(* IEC 61131-3 sources: STAR-PLC-Agent/results/raw/codex_matrix_resume_20261114/codex_deepseek/PUB002/functional/attempt_0001, 1 file *)

(* ---- test_program.st ---- *)
PROGRAM PLC_PRG
VAR
 BenchStep : UDINT := 0;
 BenchCalls : UDINT := 0;
 BenchDone : BOOL := FALSE;
 BenchUut0 : FB_Task;
 BenchUut1 : FB_Task;
 BenchUut2 : FB_Task;
 BenchUut3 : FB_Task;
 BenchUut4 : FB_Task;
 BenchUut5 : FB_Task;
 BenchUut6 : FB_Task;
 TraceIn_value : ARRAY[0..38] OF DWORD;
 TraceOut_hasChanged : ARRAY[0..38] OF BOOL;
 TraceOut_hasRisingEdges : ARRAY[0..38] OF BOOL;
 TraceOut_risingBits : ARRAY[0..38] OF DWORD;
 TraceOut_noOfRisingBits : ARRAY[0..38] OF USINT;
 TraceOut_hasFallingEdges : ARRAY[0..38] OF BOOL;
 TraceOut_fallingBits : ARRAY[0..38] OF DWORD;
 TraceOut_noOfFallingBits : ARRAY[0..38] OF USINT;
END_VAR

IF NOT BenchDone THEN
 CASE BenchStep OF
 0:
   BenchUut0.value := DWORD#0;
   TraceIn_value[0] := BenchUut0.value;
   BenchUut0();
   TraceOut_hasChanged[0] := BenchUut0.hasChanged;
   TraceOut_hasRisingEdges[0] := BenchUut0.hasRisingEdges;
   TraceOut_risingBits[0] := BenchUut0.risingBits;
   TraceOut_noOfRisingBits[0] := BenchUut0.noOfRisingBits;
   TraceOut_hasFallingEdges[0] := BenchUut0.hasFallingEdges;
   TraceOut_fallingBits[0] := BenchUut0.fallingBits;
   TraceOut_noOfFallingBits[0] := BenchUut0.noOfFallingBits;
   BenchCalls := BenchCalls + 1;
 1:
   BenchUut0.value := DWORD#1;
   TraceIn_value[1] := BenchUut0.value;
   BenchUut0();
   TraceOut_hasChanged[1] := BenchUut0.hasChanged;
   TraceOut_hasRisingEdges[1] := BenchUut0.hasRisingEdges;
   TraceOut_risingBits[1] := BenchUut0.risingBits;
   TraceOut_noOfRisingBits[1] := BenchUut0.noOfRisingBits;
   TraceOut_hasFallingEdges[1] := BenchUut0.hasFallingEdges;
   TraceOut_fallingBits[1] := BenchUut0.fallingBits;
   TraceOut_noOfFallingBits[1] := BenchUut0.noOfFallingBits;
   BenchCalls := BenchCalls + 1;
 2:
   BenchUut0.value := DWORD#1;
   TraceIn_value[2] := BenchUut0.value;
   BenchUut0();
   TraceOut_hasChanged[2] := BenchUut0.hasChanged;
   TraceOut_hasRisingEdges[2] := BenchUut0.hasRisingEdges;
   TraceOut_risingBits[2] := BenchUut0.risingBits;
   TraceOut_noOfRisingBits[2] := BenchUut0.noOfRisingBits;
   TraceOut_hasFallingEdges[2] := BenchUut0.hasFallingEdges;
   TraceOut_fallingBits[2] := BenchUut0.fallingBits;
   TraceOut_noOfFallingBits[2] := BenchUut0.noOfFallingBits;
   BenchCalls := BenchCalls + 1;
 3:
   BenchUut0.value := DWORD#3;
   TraceIn_value[3] := BenchUut0.value;
   BenchUut0();
   TraceOut_hasChanged[3] := BenchUut0.hasChanged;
   TraceOut_hasRisingEdges[3] := BenchUut0.hasRisingEdges;
   TraceOut_risingBits[3] := BenchUut0.risingBits;
   TraceOut_noOfRisingBits[3] := BenchUut0.noOfRisingBits;
   TraceOut_hasFallingEdges[3] := BenchUut0.hasFallingEdges;
   TraceOut_fallingBits[3] := BenchUut0.fallingBits;
   TraceOut_noOfFallingBits[3] := BenchUut0.noOfFallingBits;
   BenchCalls := BenchCalls + 1;
 4:
   BenchUut0.value := DWORD#2;
   TraceIn_value[4] := BenchUut0.value;
   BenchUut0();
   TraceOut_hasChanged[4] := BenchUut0.hasChanged;
   TraceOut_hasRisingEdges[4] := BenchUut0.hasRisingEdges;
   TraceOut_risingBits[4] := BenchUut0.risingBits;
   TraceOut_noOfRisingBits[4] := BenchUut0.noOfRisingBits;
   TraceOut_hasFallingEdges[4] := BenchUut0.hasFallingEdges;
   TraceOut_fallingBits[4] := BenchUut0.fallingBits;
   TraceOut_noOfFallingBits[4] := BenchUut0.noOfFallingBits;
   BenchCalls := BenchCalls + 1;
 5:
   BenchUut0.value := DWORD#0;
   TraceIn_value[5] := BenchUut0.value;
   BenchUut0();
   TraceOut_hasChanged[5] := BenchUut0.hasChanged;
   TraceOut_hasRisingEdges[5] := BenchUut0.hasRisingEdges;
   TraceOut_risingBits[5] := BenchUut0.risingBits;
   TraceOut_noOfRisingBits[5] := BenchUut0.noOfRisingBits;
   TraceOut_hasFallingEdges[5] := BenchUut0.hasFallingEdges;
   TraceOut_fallingBits[5] := BenchUut0.fallingBits;
   TraceOut_noOfFallingBits[5] := BenchUut0.noOfFallingBits;
   BenchCalls := BenchCalls + 1;
 6:
   BenchUut0.value := DWORD#4294967295;
   TraceIn_value[6] := BenchUut0.value;
   BenchUut0();
   TraceOut_hasChanged[6] := BenchUut0.hasChanged;
   TraceOut_hasRisingEdges[6] := BenchUut0.hasRisingEdges;
   TraceOut_risingBits[6] := BenchUut0.risingBits;
   TraceOut_noOfRisingBits[6] := BenchUut0.noOfRisingBits;
   TraceOut_hasFallingEdges[6] := BenchUut0.hasFallingEdges;
   TraceOut_fallingBits[6] := BenchUut0.fallingBits;
   TraceOut_noOfFallingBits[6] := BenchUut0.noOfFallingBits;
   BenchCalls := BenchCalls + 1;
 7:
   BenchUut0.value := DWORD#0;
   TraceIn_value[7] := BenchUut0.value;
   BenchUut0();
   TraceOut_hasChanged[7] := BenchUut0.hasChanged;
   TraceOut_hasRisingEdges[7] := BenchUut0.hasRisingEdges;
   TraceOut_risingBits[7] := BenchUut0.risingBits;
   TraceOut_noOfRisingBits[7] := BenchUut0.noOfRisingBits;
   TraceOut_hasFallingEdges[7] := BenchUut0.hasFallingEdges;
   TraceOut_fallingBits[7] := BenchUut0.fallingBits;
   TraceOut_noOfFallingBits[7] := BenchUut0.noOfFallingBits;
   BenchCalls := BenchCalls + 1;
 8:
   BenchUut0.value := DWORD#2147483648;
   TraceIn_value[8] := BenchUut0.value;
   BenchUut0();
   TraceOut_hasChanged[8] := BenchUut0.hasChanged;
   TraceOut_hasRisingEdges[8] := BenchUut0.hasRisingEdges;
   TraceOut_risingBits[8] := BenchUut0.risingBits;
   TraceOut_noOfRisingBits[8] := BenchUut0.noOfRisingBits;
   TraceOut_hasFallingEdges[8] := BenchUut0.hasFallingEdges;
   TraceOut_fallingBits[8] := BenchUut0.fallingBits;
   TraceOut_noOfFallingBits[8] := BenchUut0.noOfFallingBits;
   BenchCalls := BenchCalls + 1;
 9:
   BenchUut0.value := DWORD#2147483647;
   TraceIn_value[9] := BenchUut0.value;
   BenchUut0();
   TraceOut_hasChanged[9] := BenchUut0.hasChanged;
   TraceOut_hasRisingEdges[9] := BenchUut0.hasRisingEdges;
   TraceOut_risingBits[9] := BenchUut0.risingBits;
   TraceOut_noOfRisingBits[9] := BenchUut0.noOfRisingBits;
   TraceOut_hasFallingEdges[9] := BenchUut0.hasFallingEdges;
   TraceOut_fallingBits[9] := BenchUut0.fallingBits;
   TraceOut_noOfFallingBits[9] := BenchUut0.noOfFallingBits;
   BenchCalls := BenchCalls + 1;
 10:
   BenchUut1.value := DWORD#4294967295;
   TraceIn_value[10] := BenchUut1.value;
   BenchUut1();
   TraceOut_hasChanged[10] := BenchUut1.hasChanged;
   TraceOut_hasRisingEdges[10] := BenchUut1.hasRisingEdges;
   TraceOut_risingBits[10] := BenchUut1.risingBits;
   TraceOut_noOfRisingBits[10] := BenchUut1.noOfRisingBits;
   TraceOut_hasFallingEdges[10] := BenchUut1.hasFallingEdges;
   TraceOut_fallingBits[10] := BenchUut1.fallingBits;
   TraceOut_noOfFallingBits[10] := BenchUut1.noOfFallingBits;
   BenchCalls := BenchCalls + 1;
 11:
   BenchUut1.value := DWORD#4294967295;
   TraceIn_value[11] := BenchUut1.value;
   BenchUut1();
   TraceOut_hasChanged[11] := BenchUut1.hasChanged;
   TraceOut_hasRisingEdges[11] := BenchUut1.hasRisingEdges;
   TraceOut_risingBits[11] := BenchUut1.risingBits;
   TraceOut_noOfRisingBits[11] := BenchUut1.noOfRisingBits;
   TraceOut_hasFallingEdges[11] := BenchUut1.hasFallingEdges;
   TraceOut_fallingBits[11] := BenchUut1.fallingBits;
   TraceOut_noOfFallingBits[11] := BenchUut1.noOfFallingBits;
   BenchCalls := BenchCalls + 1;
 12:
   BenchUut2.value := DWORD#2863311530;
   TraceIn_value[12] := BenchUut2.value;
   BenchUut2();
   TraceOut_hasChanged[12] := BenchUut2.hasChanged;
   TraceOut_hasRisingEdges[12] := BenchUut2.hasRisingEdges;
   TraceOut_risingBits[12] := BenchUut2.risingBits;
   TraceOut_noOfRisingBits[12] := BenchUut2.noOfRisingBits;
   TraceOut_hasFallingEdges[12] := BenchUut2.hasFallingEdges;
   TraceOut_fallingBits[12] := BenchUut2.fallingBits;
   TraceOut_noOfFallingBits[12] := BenchUut2.noOfFallingBits;
   BenchCalls := BenchCalls + 1;
 13:
   BenchUut2.value := DWORD#1431655765;
   TraceIn_value[13] := BenchUut2.value;
   BenchUut2();
   TraceOut_hasChanged[13] := BenchUut2.hasChanged;
   TraceOut_hasRisingEdges[13] := BenchUut2.hasRisingEdges;
   TraceOut_risingBits[13] := BenchUut2.risingBits;
   TraceOut_noOfRisingBits[13] := BenchUut2.noOfRisingBits;
   TraceOut_hasFallingEdges[13] := BenchUut2.hasFallingEdges;
   TraceOut_fallingBits[13] := BenchUut2.fallingBits;
   TraceOut_noOfFallingBits[13] := BenchUut2.noOfFallingBits;
   BenchCalls := BenchCalls + 1;
 14:
   BenchUut3.value := DWORD#983295;
   TraceIn_value[14] := BenchUut3.value;
   BenchUut3();
   TraceOut_hasChanged[14] := BenchUut3.hasChanged;
   TraceOut_hasRisingEdges[14] := BenchUut3.hasRisingEdges;
   TraceOut_risingBits[14] := BenchUut3.risingBits;
   TraceOut_noOfRisingBits[14] := BenchUut3.noOfRisingBits;
   TraceOut_hasFallingEdges[14] := BenchUut3.hasFallingEdges;
   TraceOut_fallingBits[14] := BenchUut3.fallingBits;
   TraceOut_noOfFallingBits[14] := BenchUut3.noOfFallingBits;
   BenchCalls := BenchCalls + 1;
 15:
   BenchUut3.value := DWORD#16715520;
   TraceIn_value[15] := BenchUut3.value;
   BenchUut3();
   TraceOut_hasChanged[15] := BenchUut3.hasChanged;
   TraceOut_hasRisingEdges[15] := BenchUut3.hasRisingEdges;
   TraceOut_risingBits[15] := BenchUut3.risingBits;
   TraceOut_noOfRisingBits[15] := BenchUut3.noOfRisingBits;
   TraceOut_hasFallingEdges[15] := BenchUut3.hasFallingEdges;
   TraceOut_fallingBits[15] := BenchUut3.fallingBits;
   TraceOut_noOfFallingBits[15] := BenchUut3.noOfFallingBits;
   BenchCalls := BenchCalls + 1;
 16:
   BenchUut3.value := DWORD#16715520;
   TraceIn_value[16] := BenchUut3.value;
   BenchUut3();
   TraceOut_hasChanged[16] := BenchUut3.hasChanged;
   TraceOut_hasRisingEdges[16] := BenchUut3.hasRisingEdges;
   TraceOut_risingBits[16] := BenchUut3.risingBits;
   TraceOut_noOfRisingBits[16] := BenchUut3.noOfRisingBits;
   TraceOut_hasFallingEdges[16] := BenchUut3.hasFallingEdges;
   TraceOut_fallingBits[16] := BenchUut3.fallingBits;
   TraceOut_noOfFallingBits[16] := BenchUut3.noOfFallingBits;
   BenchCalls := BenchCalls + 1;
 17:
   BenchUut3.value := DWORD#4294967295;
   TraceIn_value[17] := BenchUut3.value;
   BenchUut3();
   TraceOut_hasChanged[17] := BenchUut3.hasChanged;
   TraceOut_hasRisingEdges[17] := BenchUut3.hasRisingEdges;
   TraceOut_risingBits[17] := BenchUut3.risingBits;
   TraceOut_noOfRisingBits[17] := BenchUut3.noOfRisingBits;
   TraceOut_hasFallingEdges[17] := BenchUut3.hasFallingEdges;
   TraceOut_fallingBits[17] := BenchUut3.fallingBits;
   TraceOut_noOfFallingBits[17] := BenchUut3.noOfFallingBits;
   BenchCalls := BenchCalls + 1;
 18:
   BenchUut3.value := DWORD#2147483649;
   TraceIn_value[18] := BenchUut3.value;
   BenchUut3();
   TraceOut_hasChanged[18] := BenchUut3.hasChanged;
   TraceOut_hasRisingEdges[18] := BenchUut3.hasRisingEdges;
   TraceOut_risingBits[18] := BenchUut3.risingBits;
   TraceOut_noOfRisingBits[18] := BenchUut3.noOfRisingBits;
   TraceOut_hasFallingEdges[18] := BenchUut3.hasFallingEdges;
   TraceOut_fallingBits[18] := BenchUut3.fallingBits;
   TraceOut_noOfFallingBits[18] := BenchUut3.noOfFallingBits;
   BenchCalls := BenchCalls + 1;
 19:
   BenchUut3.value := DWORD#0;
   TraceIn_value[19] := BenchUut3.value;
   BenchUut3();
   TraceOut_hasChanged[19] := BenchUut3.hasChanged;
   TraceOut_hasRisingEdges[19] := BenchUut3.hasRisingEdges;
   TraceOut_risingBits[19] := BenchUut3.risingBits;
   TraceOut_noOfRisingBits[19] := BenchUut3.noOfRisingBits;
   TraceOut_hasFallingEdges[19] := BenchUut3.hasFallingEdges;
   TraceOut_fallingBits[19] := BenchUut3.fallingBits;
   TraceOut_noOfFallingBits[19] := BenchUut3.noOfFallingBits;
   BenchCalls := BenchCalls + 1;
 20:
   BenchUut4.value := DWORD#0;
   TraceIn_value[20] := BenchUut4.value;
   BenchUut4();
   TraceOut_hasChanged[20] := BenchUut4.hasChanged;
   TraceOut_hasRisingEdges[20] := BenchUut4.hasRisingEdges;
   TraceOut_risingBits[20] := BenchUut4.risingBits;
   TraceOut_noOfRisingBits[20] := BenchUut4.noOfRisingBits;
   TraceOut_hasFallingEdges[20] := BenchUut4.hasFallingEdges;
   TraceOut_fallingBits[20] := BenchUut4.fallingBits;
   TraceOut_noOfFallingBits[20] := BenchUut4.noOfFallingBits;
   BenchCalls := BenchCalls + 1;
 21:
   BenchUut4.value := DWORD#2;
   TraceIn_value[21] := BenchUut4.value;
   BenchUut4();
   TraceOut_hasChanged[21] := BenchUut4.hasChanged;
   TraceOut_hasRisingEdges[21] := BenchUut4.hasRisingEdges;
   TraceOut_risingBits[21] := BenchUut4.risingBits;
   TraceOut_noOfRisingBits[21] := BenchUut4.noOfRisingBits;
   TraceOut_hasFallingEdges[21] := BenchUut4.hasFallingEdges;
   TraceOut_fallingBits[21] := BenchUut4.fallingBits;
   TraceOut_noOfFallingBits[21] := BenchUut4.noOfFallingBits;
   BenchCalls := BenchCalls + 1;
 22:
   BenchUut4.value := DWORD#2;
   TraceIn_value[22] := BenchUut4.value;
   BenchUut4();
   TraceOut_hasChanged[22] := BenchUut4.hasChanged;
   TraceOut_hasRisingEdges[22] := BenchUut4.hasRisingEdges;
   TraceOut_risingBits[22] := BenchUut4.risingBits;
   TraceOut_noOfRisingBits[22] := BenchUut4.noOfRisingBits;
   TraceOut_hasFallingEdges[22] := BenchUut4.hasFallingEdges;
   TraceOut_fallingBits[22] := BenchUut4.fallingBits;
   TraceOut_noOfFallingBits[22] := BenchUut4.noOfFallingBits;
   BenchCalls := BenchCalls + 1;
 23:
   BenchUut4.value := DWORD#8;
   TraceIn_value[23] := BenchUut4.value;
   BenchUut4();
   TraceOut_hasChanged[23] := BenchUut4.hasChanged;
   TraceOut_hasRisingEdges[23] := BenchUut4.hasRisingEdges;
   TraceOut_risingBits[23] := BenchUut4.risingBits;
   TraceOut_noOfRisingBits[23] := BenchUut4.noOfRisingBits;
   TraceOut_hasFallingEdges[23] := BenchUut4.hasFallingEdges;
   TraceOut_fallingBits[23] := BenchUut4.fallingBits;
   TraceOut_noOfFallingBits[23] := BenchUut4.noOfFallingBits;
   BenchCalls := BenchCalls + 1;
 24:
   BenchUut4.value := DWORD#8;
   TraceIn_value[24] := BenchUut4.value;
   BenchUut4();
   TraceOut_hasChanged[24] := BenchUut4.hasChanged;
   TraceOut_hasRisingEdges[24] := BenchUut4.hasRisingEdges;
   TraceOut_risingBits[24] := BenchUut4.risingBits;
   TraceOut_noOfRisingBits[24] := BenchUut4.noOfRisingBits;
   TraceOut_hasFallingEdges[24] := BenchUut4.hasFallingEdges;
   TraceOut_fallingBits[24] := BenchUut4.fallingBits;
   TraceOut_noOfFallingBits[24] := BenchUut4.noOfFallingBits;
   BenchCalls := BenchCalls + 1;
 25:
   BenchUut4.value := DWORD#10;
   TraceIn_value[25] := BenchUut4.value;
   BenchUut4();
   TraceOut_hasChanged[25] := BenchUut4.hasChanged;
   TraceOut_hasRisingEdges[25] := BenchUut4.hasRisingEdges;
   TraceOut_risingBits[25] := BenchUut4.risingBits;
   TraceOut_noOfRisingBits[25] := BenchUut4.noOfRisingBits;
   TraceOut_hasFallingEdges[25] := BenchUut4.hasFallingEdges;
   TraceOut_fallingBits[25] := BenchUut4.fallingBits;
   TraceOut_noOfFallingBits[25] := BenchUut4.noOfFallingBits;
   BenchCalls := BenchCalls + 1;
 26:
   BenchUut4.value := DWORD#0;
   TraceIn_value[26] := BenchUut4.value;
   BenchUut4();
   TraceOut_hasChanged[26] := BenchUut4.hasChanged;
   TraceOut_hasRisingEdges[26] := BenchUut4.hasRisingEdges;
   TraceOut_risingBits[26] := BenchUut4.risingBits;
   TraceOut_noOfRisingBits[26] := BenchUut4.noOfRisingBits;
   TraceOut_hasFallingEdges[26] := BenchUut4.hasFallingEdges;
   TraceOut_fallingBits[26] := BenchUut4.fallingBits;
   TraceOut_noOfFallingBits[26] := BenchUut4.noOfFallingBits;
   BenchCalls := BenchCalls + 1;
 27:
   BenchUut4.value := DWORD#0;
   TraceIn_value[27] := BenchUut4.value;
   BenchUut4();
   TraceOut_hasChanged[27] := BenchUut4.hasChanged;
   TraceOut_hasRisingEdges[27] := BenchUut4.hasRisingEdges;
   TraceOut_risingBits[27] := BenchUut4.risingBits;
   TraceOut_noOfRisingBits[27] := BenchUut4.noOfRisingBits;
   TraceOut_hasFallingEdges[27] := BenchUut4.hasFallingEdges;
   TraceOut_fallingBits[27] := BenchUut4.fallingBits;
   TraceOut_noOfFallingBits[27] := BenchUut4.noOfFallingBits;
   BenchCalls := BenchCalls + 1;
 28:
   BenchUut5.value := DWORD#0;
   TraceIn_value[28] := BenchUut5.value;
   BenchUut5();
   TraceOut_hasChanged[28] := BenchUut5.hasChanged;
   TraceOut_hasRisingEdges[28] := BenchUut5.hasRisingEdges;
   TraceOut_risingBits[28] := BenchUut5.risingBits;
   TraceOut_noOfRisingBits[28] := BenchUut5.noOfRisingBits;
   TraceOut_hasFallingEdges[28] := BenchUut5.hasFallingEdges;
   TraceOut_fallingBits[28] := BenchUut5.fallingBits;
   TraceOut_noOfFallingBits[28] := BenchUut5.noOfFallingBits;
   BenchCalls := BenchCalls + 1;
 29:
   BenchUut5.value := DWORD#4294901760;
   TraceIn_value[29] := BenchUut5.value;
   BenchUut5();
   TraceOut_hasChanged[29] := BenchUut5.hasChanged;
   TraceOut_hasRisingEdges[29] := BenchUut5.hasRisingEdges;
   TraceOut_risingBits[29] := BenchUut5.risingBits;
   TraceOut_noOfRisingBits[29] := BenchUut5.noOfRisingBits;
   TraceOut_hasFallingEdges[29] := BenchUut5.hasFallingEdges;
   TraceOut_fallingBits[29] := BenchUut5.fallingBits;
   TraceOut_noOfFallingBits[29] := BenchUut5.noOfFallingBits;
   BenchCalls := BenchCalls + 1;
 30:
   BenchUut5.value := DWORD#65535;
   TraceIn_value[30] := BenchUut5.value;
   BenchUut5();
   TraceOut_hasChanged[30] := BenchUut5.hasChanged;
   TraceOut_hasRisingEdges[30] := BenchUut5.hasRisingEdges;
   TraceOut_risingBits[30] := BenchUut5.risingBits;
   TraceOut_noOfRisingBits[30] := BenchUut5.noOfRisingBits;
   TraceOut_hasFallingEdges[30] := BenchUut5.hasFallingEdges;
   TraceOut_fallingBits[30] := BenchUut5.fallingBits;
   TraceOut_noOfFallingBits[30] := BenchUut5.noOfFallingBits;
   BenchCalls := BenchCalls + 1;
 31:
   BenchUut5.value := DWORD#2147483649;
   TraceIn_value[31] := BenchUut5.value;
   BenchUut5();
   TraceOut_hasChanged[31] := BenchUut5.hasChanged;
   TraceOut_hasRisingEdges[31] := BenchUut5.hasRisingEdges;
   TraceOut_risingBits[31] := BenchUut5.risingBits;
   TraceOut_noOfRisingBits[31] := BenchUut5.noOfRisingBits;
   TraceOut_hasFallingEdges[31] := BenchUut5.hasFallingEdges;
   TraceOut_fallingBits[31] := BenchUut5.fallingBits;
   TraceOut_noOfFallingBits[31] := BenchUut5.noOfFallingBits;
   BenchCalls := BenchCalls + 1;
 32:
   BenchUut5.value := DWORD#2147483646;
   TraceIn_value[32] := BenchUut5.value;
   BenchUut5();
   TraceOut_hasChanged[32] := BenchUut5.hasChanged;
   TraceOut_hasRisingEdges[32] := BenchUut5.hasRisingEdges;
   TraceOut_risingBits[32] := BenchUut5.risingBits;
   TraceOut_noOfRisingBits[32] := BenchUut5.noOfRisingBits;
   TraceOut_hasFallingEdges[32] := BenchUut5.hasFallingEdges;
   TraceOut_fallingBits[32] := BenchUut5.fallingBits;
   TraceOut_noOfFallingBits[32] := BenchUut5.noOfFallingBits;
   BenchCalls := BenchCalls + 1;
 33:
   BenchUut5.value := DWORD#2147483646;
   TraceIn_value[33] := BenchUut5.value;
   BenchUut5();
   TraceOut_hasChanged[33] := BenchUut5.hasChanged;
   TraceOut_hasRisingEdges[33] := BenchUut5.hasRisingEdges;
   TraceOut_risingBits[33] := BenchUut5.risingBits;
   TraceOut_noOfRisingBits[33] := BenchUut5.noOfRisingBits;
   TraceOut_hasFallingEdges[33] := BenchUut5.hasFallingEdges;
   TraceOut_fallingBits[33] := BenchUut5.fallingBits;
   TraceOut_noOfFallingBits[33] := BenchUut5.noOfFallingBits;
   BenchCalls := BenchCalls + 1;
 34:
   BenchUut6.value := DWORD#4294967295;
   TraceIn_value[34] := BenchUut6.value;
   BenchUut6();
   TraceOut_hasChanged[34] := BenchUut6.hasChanged;
   TraceOut_hasRisingEdges[34] := BenchUut6.hasRisingEdges;
   TraceOut_risingBits[34] := BenchUut6.risingBits;
   TraceOut_noOfRisingBits[34] := BenchUut6.noOfRisingBits;
   TraceOut_hasFallingEdges[34] := BenchUut6.hasFallingEdges;
   TraceOut_fallingBits[34] := BenchUut6.fallingBits;
   TraceOut_noOfFallingBits[34] := BenchUut6.noOfFallingBits;
   BenchCalls := BenchCalls + 1;
 35:
   BenchUut6.value := DWORD#2863311530;
   TraceIn_value[35] := BenchUut6.value;
   BenchUut6();
   TraceOut_hasChanged[35] := BenchUut6.hasChanged;
   TraceOut_hasRisingEdges[35] := BenchUut6.hasRisingEdges;
   TraceOut_risingBits[35] := BenchUut6.risingBits;
   TraceOut_noOfRisingBits[35] := BenchUut6.noOfRisingBits;
   TraceOut_hasFallingEdges[35] := BenchUut6.hasFallingEdges;
   TraceOut_fallingBits[35] := BenchUut6.fallingBits;
   TraceOut_noOfFallingBits[35] := BenchUut6.noOfFallingBits;
   BenchCalls := BenchCalls + 1;
 36:
   BenchUut6.value := DWORD#1431655765;
   TraceIn_value[36] := BenchUut6.value;
   BenchUut6();
   TraceOut_hasChanged[36] := BenchUut6.hasChanged;
   TraceOut_hasRisingEdges[36] := BenchUut6.hasRisingEdges;
   TraceOut_risingBits[36] := BenchUut6.risingBits;
   TraceOut_noOfRisingBits[36] := BenchUut6.noOfRisingBits;
   TraceOut_hasFallingEdges[36] := BenchUut6.hasFallingEdges;
   TraceOut_fallingBits[36] := BenchUut6.fallingBits;
   TraceOut_noOfFallingBits[36] := BenchUut6.noOfFallingBits;
   BenchCalls := BenchCalls + 1;
 37:
   BenchUut6.value := DWORD#0;
   TraceIn_value[37] := BenchUut6.value;
   BenchUut6();
   TraceOut_hasChanged[37] := BenchUut6.hasChanged;
   TraceOut_hasRisingEdges[37] := BenchUut6.hasRisingEdges;
   TraceOut_risingBits[37] := BenchUut6.risingBits;
   TraceOut_noOfRisingBits[37] := BenchUut6.noOfRisingBits;
   TraceOut_hasFallingEdges[37] := BenchUut6.hasFallingEdges;
   TraceOut_fallingBits[37] := BenchUut6.fallingBits;
   TraceOut_noOfFallingBits[37] := BenchUut6.noOfFallingBits;
   BenchCalls := BenchCalls + 1;
 38:
   BenchUut6.value := DWORD#1;
   TraceIn_value[38] := BenchUut6.value;
   BenchUut6();
   TraceOut_hasChanged[38] := BenchUut6.hasChanged;
   TraceOut_hasRisingEdges[38] := BenchUut6.hasRisingEdges;
   TraceOut_risingBits[38] := BenchUut6.risingBits;
   TraceOut_noOfRisingBits[38] := BenchUut6.noOfRisingBits;
   TraceOut_hasFallingEdges[38] := BenchUut6.hasFallingEdges;
   TraceOut_fallingBits[38] := BenchUut6.fallingBits;
   TraceOut_noOfFallingBits[38] := BenchUut6.noOfFallingBits;
   BenchCalls := BenchCalls + 1;
 END_CASE;
 BenchStep := BenchStep + 1;
 IF BenchStep >= 39 THEN BenchDone := TRUE; END_IF;
END_IF;
END_PROGRAM
